(* IEC 61131-3 sources: plc-vscode/tests/st/all/trust-platform/examples/plcopen_motion_single_axis_benchmarks/runtime_floor/src, 2 files *)

(* ---- Globals.st ---- *)
VAR_GLOBAL
    g_motion_bench_cycles : UDINT;
    g_motion_bench_completed_sequences : UDINT;
    g_motion_bench_last_error : WORD;
    g_motion_bench_power_on : BOOL;
    g_motion_bench_is_homed : BOOL;
    g_motion_bench_last_position : REAL;
    g_motion_bench_last_velocity : REAL;
    g_motion_bench_current_step : UINT;
END_VAR

(* ---- Main.st ---- *)
PROGRAM Main
g_motion_bench_cycles := g_motion_bench_cycles + UDINT#1;
g_motion_bench_completed_sequences := g_motion_bench_cycles;
g_motion_bench_last_error := WORD#16#0000;
g_motion_bench_power_on := FALSE;
g_motion_bench_is_homed := FALSE;
g_motion_bench_last_position := REAL#0.0;
g_motion_bench_last_velocity := REAL#0.0;
g_motion_bench_current_step := UINT#1;
END_PROGRAM
